// TIA Portal V20 export
// export: Created 2026-10-20T12:46:06.1060455Z, ExportSetting WithDefaults, DisplayName Totally Integrated Automation Portal, DisplayVersion V20 Update 6, DisplayName TIA Portal Openness, DisplayVersion V20 Update 6, DisplayName TIA Portal Version Control Interface, DisplayVersion V20 Update 6, DisplayName SINAMICS Startdrive Advanced, DisplayVersion V20 SP1, DisplayName SINAMICS Startdrive G130, G150, S120, S150, SINAMICS MV, G220, S200, S210, DisplayVersion V20 SP1, DisplayName SINAMICS Startdrive G110M, G120, G120C, G120D, G120P, G115D, DisplayVersion V20 SP1, DisplayName STEP 7 Professional, DisplayVersion V20 Update 6, DisplayName STEP 7 Safety, DisplayVersion V20 Update 2, DisplayName WinCC Basic/Comfort/Advanced, DisplayVersion V20 Update 6, DisplayName WinCC Unified, DisplayVersion V20 Update 6
DATA_BLOCK "PopUps_DB"   // DB38
{ S7_Optimized_Access := 'TRUE' }
VERSION : 0.1
// stored: AutoNumber false, DBAccessibleFromOPCUA true, IsOnlyStoredInLoadMemory false, IsRetainMemResEnabled false, IsWriteProtectedInAS false, MemoryReserve 100
   VAR
      Buffer_Cnv_Settings_1 : "Buffer_Cnv_Settings";
      Buffer_Cnv_Settings_2 { S7_SetPoint := 'True'} : "Buffer_Cnv_Settings";
      ECnv_Settings { S7_SetPoint := 'True'} : "ECnv_Settings";
      VTD_Settings { S7_SetPoint := 'True'} : "VTD_Settings";
      Shuttle_MQTT_Settings { S7_SetPoint := 'True'} : "MQTT_Settings";
      Sick_Lector_Reseult : String;
   END_VAR
BEGIN
END_DATA_BLOCK
